(* IEC 61131-3 sources: plc-st-coding-agent/progress/evidence/f14_v14_remaining_20261113/jobs/custom_minimax-m27 (part 2) *)

(* ---- public-hard-03.raw_candidate_01.st ---- *)
FUNCTION_BLOCK FB_RecipeManager
VAR_INPUT
    addRecipe      : BOOL;
    deleteRecipe   : BOOL;
    modifyRecipe   : BOOL;
    queryRecipe    : BOOL;
    recipeIn       : ST_Recipe;
END_VAR

VAR_OUTPUT
    recipeAdded        : BOOL;
    recipeDeleted      : BOOL;
    recipeModified     : BOOL;
    recipeQueryResult  : ST_Recipe;
    error              : BOOL;
    status             : WORD;
END_VAR

VAR_IN_OUT
    recipe : ARRAY[1..10] OF ST_Recipe;
END_VAR

VAR
    tmp_foundIndex : INT;
    tmp_emptyIndex : INT;
    tmp_i          : INT;
END_VAR

(*
ENGINEERING_CONTRACT
===================
Operation sequencing (PUB001-PUB005, PUB007-PUB012):
- Commands evaluated in priority order: DELETE > ADD > MODIFY > QUERY when multiple asserted.
- All success pulses are same-scan; no retention across scans.

Query (PUB008):
  Activation:    queryRecipe rising edge or held high during scan.
  Retention:     recipeQueryResult valid until next scan or successful QUERY.
  Reset:         error and status cleared at start of scan.
  Error codes:   16#8001 = recipe not found.
  Units:         Status WORD error code.

Add (PUB009):
  Activation:    addRecipe rising edge or held high.
  Retention:     Stored in smallest-index empty slot; persists until delete.
  Reset:         None (persistent storage).
  Error codes:   16#8002 = duplicate ID; 16#8003 = database full.
  Same-scan:     Duplicate check before empty-slot check.

Delete (PUB010):
  Activation:    deleteRecipe rising edge or held high.
  Retention:     recipeID forced to 0 (empty slot marker).
  Reset:         Implicit (setting ID to 0 removes it).
  Error codes:   16#8004 = recipe not found.

Modify (PUB011-PUB012):
  Activation:    modifyRecipe rising edge or held high.
  Retention:     Full recipe replacement at found slot.
  Reset:         None.
  Error codes:   16#8005 = recipe not found.
*)

(* CONTRACT_RULES [] *)

tmp_foundIndex := 0;
tmp_emptyIndex := 0;
error := FALSE;
status := 16#0;
recipeAdded := FALSE;
recipeDeleted := FALSE;
recipeModified := FALSE;

IF deleteRecipe THEN
    tmp_foundIndex := 0;
    FOR tmp_i := 1 TO 10 DO
        IF recipe[tmp_i].recipeID <> 0 AND recipe[tmp_i].recipeID = recipeIn.recipeID THEN
            tmp_foundIndex := tmp_i;
            EXIT;
        END_IF
    END_FOR;

    IF tmp_foundIndex = 0 THEN
        error := TRUE;
        status := 16#8004;
    ELSE
        recipe[tmp_foundIndex].recipeID := 0;
        recipeDeleted := TRUE;
    END_IF;

ELSIF addRecipe THEN
    tmp_foundIndex := 0;
    tmp_emptyIndex := 0;

    FOR tmp_i := 1 TO 10 DO
        IF recipe[tmp_i].recipeID <> 0 AND recipe[tmp_i].recipeID = recipeIn.recipeID THEN
            tmp_foundIndex := tmp_i;
            EXIT;
        END_IF
    END_FOR;

    IF tmp_foundIndex <> 0 THEN
        error := TRUE;
        status := 16#8002;
    ELSE
        FOR tmp_i := 1 TO 10 DO
            IF recipe[tmp_i].recipeID = 0 AND tmp_emptyIndex = 0 THEN
                tmp_emptyIndex := tmp_i;
                EXIT;
            END_IF
        END_FOR;

        IF tmp_emptyIndex = 0 THEN
            error := TRUE;
            status := 16#8003;
        ELSE
            recipe[tmp_emptyIndex] := recipeIn;
            recipeAdded := TRUE;
        END_IF;
    END_IF;

ELSIF modifyRecipe THEN
    tmp_foundIndex := 0;
    FOR tmp_i := 1 TO 10 DO
        IF recipe[tmp_i].recipeID <> 0 AND recipe[tmp_i].recipeID = recipeIn.recipeID THEN
            tmp_foundIndex := tmp_i;
            EXIT;
        END_IF
    END_FOR;

    IF tmp_foundIndex = 0 THEN
        error := TRUE;
        status := 16#8005;
    ELSE
        recipe[tmp_foundIndex] := recipeIn;
        recipeModified := TRUE;
    END_IF;

ELSIF queryRecipe THEN
    tmp_foundIndex := 0;
    FOR tmp_i := 1 TO 10 DO
        IF recipe[tmp_i].recipeID <> 0 AND recipe[tmp_i].recipeID = recipeIn.recipeID THEN
            tmp_foundIndex := tmp_i;
            EXIT;
        END_IF
    END_FOR;

    IF tmp_foundIndex = 0 THEN
        error := TRUE;
        status := 16#8001;
    ELSE
        recipeQueryResult := recipe[tmp_foundIndex];
    END_IF;
END_IF;

END_FUNCTION_BLOCK

(* ---- public-hard-03.raw_candidate_02.st ---- *)
TYPE ST_Recipe :
STRUCT
    recipeID               : INT;
    ingredientType         : INT;
    ingredientRatio        : REAL;
    productionTemperature  : REAL;
END_STRUCT
END_TYPE

FUNCTION_BLOCK FB_RecipeManager
VAR_INPUT
    addRecipe      : BOOL;
    deleteRecipe   : BOOL;
    modifyRecipe   : BOOL;
    queryRecipe    : BOOL;
    recipeIn       : ST_Recipe;
END_VAR

VAR_OUTPUT
    recipeAdded        : BOOL;
    recipeDeleted      : BOOL;
    recipeModified     : BOOL;
    recipeQueryResult  : ST_Recipe;
    error              : BOOL;
    status             : WORD;
END_VAR

VAR_IN_OUT
    recipe : ARRAY[1..10] OF ST_Recipe;
END_VAR

VAR
    tmp_foundIndex : INT;
    tmp_emptyIndex : INT;
    tmp_i          : INT;
END_VAR

(*
ENGINEERING_CONTRACT
===================
Operation sequencing (PUB001-PUB005, PUB007-PUB012):
- Commands evaluated in priority order: DELETE > ADD > MODIFY > QUERY when multiple asserted.
- All success pulses are same-scan; no retention across scans.

Query (PUB008):
  Activation:    queryRecipe rising edge or held high during scan.
  Retention:     recipeQueryResult valid until next scan or successful QUERY.
  Reset:         error and status cleared at start of scan.
  Error codes:   16#8001 = recipe not found.
  Units:         Status WORD error code.

Add (PUB009):
  Activation:    addRecipe rising edge or held high.
  Retention:     Stored in smallest-index empty slot; persists until delete.
  Reset:         None (persistent storage).
  Error codes:   16#8002 = duplicate ID; 16#8003 = database full.
  Same-scan:     Duplicate check before empty-slot check.

Delete (PUB010):
  Activation:    deleteRecipe rising edge or held high.
  Retention:     recipeID forced to 0 (empty slot marker).
  Reset:         Implicit (setting ID to 0 removes it).
  Error codes:   16#8004 = recipe not found.

Modify (PUB011-PUB012):
  Activation:    modifyRecipe rising edge or held high.
  Retention:     Full recipe replacement at found slot.
  Reset:         None.
  Error codes:   16#8005 = recipe not found.
*)

(* CONTRACT_RULES [] *)

tmp_foundIndex := 0;
tmp_emptyIndex := 0;
error := FALSE;
status := 16#0;
recipeAdded := FALSE;
recipeDeleted := FALSE;
recipeModified := FALSE;

IF deleteRecipe THEN
    tmp_foundIndex := 0;
    FOR tmp_i := 1 TO 10 DO
        IF recipe[tmp_i].recipeID <> 0 AND recipe[tmp_i].recipeID = recipeIn.recipeID THEN
            tmp_foundIndex := tmp_i;
            EXIT;
        END_IF;
    END_FOR;

    IF tmp_foundIndex = 0 THEN
        error := TRUE;
        status := 16#8004;
    ELSE
        recipe[tmp_foundIndex].recipeID := 0;
        recipeDeleted := TRUE;
    END_IF;

ELSIF addRecipe THEN
    tmp_foundIndex := 0;
    tmp_emptyIndex := 0;

    FOR tmp_i := 1 TO 10 DO
        IF recipe[tmp_i].recipeID <> 0 AND recipe[tmp_i].recipeID = recipeIn.recipeID THEN
            tmp_foundIndex := tmp_i;
            EXIT;
        END_IF;
    END_FOR;

    IF tmp_foundIndex <> 0 THEN
        error := TRUE;
        status := 16#8002;
    ELSE
        FOR tmp_i := 1 TO 10 DO
            IF recipe[tmp_i].recipeID = 0 AND tmp_emptyIndex = 0 THEN
                tmp_emptyIndex := tmp_i;
                EXIT;
            END_IF;
        END_FOR;

        IF tmp_emptyIndex = 0 THEN
            error := TRUE;
            status := 16#8003;
        ELSE
            recipe[tmp_emptyIndex] := recipeIn;
            recipeAdded := TRUE;
        END_IF;
    END_IF;

ELSIF modifyRecipe THEN
    tmp_foundIndex := 0;
    FOR tmp_i := 1 TO 10 DO
        IF recipe[tmp_i].recipeID <> 0 AND recipe[tmp_i].recipeID = recipeIn.recipeID THEN
            tmp_foundIndex := tmp_i;
            EXIT;
        END_IF;
    END_FOR;

    IF tmp_foundIndex = 0 THEN
        error := TRUE;
        status := 16#8005;
    ELSE
        recipe[tmp_foundIndex] := recipeIn;
        recipeModified := TRUE;
    END_IF;

ELSIF queryRecipe THEN
    tmp_foundIndex := 0;
    FOR tmp_i := 1 TO 10 DO
        IF recipe[tmp_i].recipeID <> 0 AND recipe[tmp_i].recipeID = recipeIn.recipeID THEN
            tmp_foundIndex := tmp_i;
            EXIT;
        END_IF;
    END_FOR;

    IF tmp_foundIndex = 0 THEN
        error := TRUE;
        status := 16#8001;
    ELSE
        recipeQueryResult := recipe[tmp_foundIndex];
    END_IF;
END_IF;

END_FUNCTION_BLOCK

(* ---- public-hard-04.candidate_01.st ---- *)
FUNCTION_BLOCK FB
VAR_INPUT
    enqueue  : BOOL;
    dequeue  : BOOL;
    reset    : BOOL;
END_VAR
VAR_OUTPUT
    elementCount : DINT := 0;
    status       : WORD := 16#0000;
END_VAR
VAR_IN_OUT
    item   : VARIANT;
    buffer : VARIANT;
END_VAR
VAR
    head          : DINT := 0;
    tail          : DINT := 0;
    enqueue_prev  : BOOL := FALSE;
    dequeue_prev  : BOOL := FALSE;
    enqueue_trig  : R_TRIG;
    dequeue_trig  : R_TRIG;
    tmp_lower     : DINT;
    tmp_upper     : DINT;
    tmp_capacity  : DINT;
    tmp_element   : DINT;
END_VAR
VAR_TEMP
    emptyArray : ARRAY[0..0] OF DINT;
END_VAR
// ENGINEERING_CONTRACT
// ─────────────────────────────────────────────────────────────────────────────
// PUB001: enqueue rising edge → write item to tail; reject if elementCount == capacity.
// PUB002: dequeue rising edge → read buffer[head] to item; reject if elementCount == 0.
// PUB003: reset TRUE → head:=0, tail:=0, elementCount:=0; no buffer overwrite.
// PUB004: elementCount output tracks live queue size (0..capacity).
// PUB005: status 16#0000=no error/idle; 16#8001=dequeue reject (empty);
//         16#8002=enqueue reject (full); 16#8003=simultaneous enqueue+dequeue.
// PUB006: buffer is caller-supplied VARIANT array; capacity = UPPER-LOWER+1.
// PUB007: item is VARIANT scalar; type must match buffer element type.
// PUB008: circular queue uses head (read index) and tail (write index) modulo capacity.
// PUB009: first invocation initializes to empty state (no prior buffer content used).
// PUB010: reset has priority over enqueue/dequeue.
// PUB011: simultaneous enqueue+dequeue is invalid usage → rejected with status 16#8003.
// ─────────────────────────────────────────────────────────────────────────────
// (* CONTRACT_RULES [] *)
// ─────────────────────────────────────────────────────────────────────────────
    // Capture rising edges for enqueue and dequeue commands
    enqueue_trig(CLK := enqueue);
    dequeue_trig(CLK := dequeue);

    // Update previous state for next scan edge detection
    enqueue_prev  := enqueue;
    dequeue_prev  := dequeue;

    // Reject simultaneous enqueue and dequeue requests
    IF enqueue AND dequeue THEN
        status := 16#8003;
        RETURN;
    END_IF;

    // Validate buffer pointer and extract array bounds
    IF __ISVALIDPTR(buffer, TO_DINT(SIZEOF(emptyArray))) THEN
        tmp_lower    := LOWER_BOUND(buffer, 1);
        tmp_upper    := UPPER_BOUND(buffer, 1);
        tmp_capacity := TO_DINT(tmp_upper - tmp_lower + 1);

        // Validate capacity is positive
        IF tmp_capacity <= 0 THEN
            status := 16#FFFF;
            RETURN;
        END_IF;

        // Type validation: ensure item type matches buffer element type
        // by reading from buffer then assigning to item (runtime type check)
        tmp_element := buffer[tmp_lower];
        tmp_element := item;

        // Execute prioritized operations
        IF reset THEN
            // PUB003: Reset clears queue state without overwriting buffer content
            head        := 0;
            tail        := 0;
            elementCount := 0;
            status      := 16#0000;
        ELSIF enqueue_trig.Q THEN
            // PUB001: Enqueue operation
            IF elementCount >= tmp_capacity THEN
                // Queue full - reject enqueue
                status := 16#8002;
            ELSE
                // Write item to tail position, advance tail circularly
                buffer[tail] := item;
                tail         := (tail + 1) MOD tmp_capacity;
                elementCount := elementCount + 1;
                status       := 16#0000;
            END_IF;
        ELSIF dequeue_trig.Q THEN
            // PUB002: Dequeue operation
            IF elementCount <= 0 THEN
                // Queue empty - reject dequeue
                status := 16#8001;
            ELSE
                // Read from head position, advance head circularly
                item        := buffer[head];
                head        := (head + 1) MOD tmp_capacity;
                elementCount := elementCount - 1;
                status       := 16#0000;
            END_IF;
        ELSE
            // No operation requested this scan
            status := 16#0000;
        END_IF;
    ELSE
        status := 16#FFFF;
    END_IF;
END_FUNCTION_BLOCK

(* ---- public-hard-04.candidate_03.st ---- *)
FUNCTION_BLOCK FB
VAR_INPUT
    enqueue  : BOOL;
    dequeue  : BOOL;
    reset    : BOOL;
END_VAR
VAR_OUTPUT
    elementCount : DINT := 0;
    status       : WORD := 16#0000;
END_VAR
VAR_IN_OUT
    item   : VARIANT;
    buffer : VARIANT;
END_VAR
VAR
    head          : DINT := 0;
    tail          : DINT := 0;
    enqueue_prev  : BOOL := FALSE;
    dequeue_prev  : BOOL := FALSE;
    enqueue_trig  : R_TRIG;
    dequeue_trig  : R_TRIG;
    tmp_lower     : DINT;
    tmp_upper     : DINT;
    tmp_capacity  : DINT;
    tmp_element   : DINT;
END_VAR
// ENGINEERING_CONTRACT
// ─────────────────────────────────────────────────────────────────────────────
// PUB001: enqueue rising edge → write item to tail; reject if elementCount == capacity.
// PUB002: dequeue rising edge → read buffer[head] to item; reject if elementCount == 0.
// PUB003: reset TRUE → head:=0, tail:=0, elementCount:=0; no buffer overwrite.
// PUB004: elementCount output tracks live queue size (0..capacity).
// PUB005: status 16#0000=no error/idle; 16#8001=dequeue reject (empty);
//         16#8002=enqueue reject (full); 16#8003=simultaneous enqueue+dequeue.
// PUB006: buffer is caller-supplied VARIANT array; capacity = UPPER-LOWER+1.
// PUB007: item is VARIANT scalar; type must match buffer element type.
// PUB008: circular queue uses head (read index) and tail (write index) modulo capacity.
// PUB009: first invocation initializes to empty state (no prior buffer content used).
// PUB010: reset has priority over enqueue/dequeue.
// PUB011: simultaneous enqueue+dequeue is invalid usage → rejected with status 16#8003.
// ─────────────────────────────────────────────────────────────────────────────
// (* CONTRACT_RULES [] *)
// ─────────────────────────────────────────────────────────────────────────────
    // Capture rising edges for enqueue and dequeue commands
    enqueue_trig(CLK := enqueue);
    dequeue_trig(CLK := dequeue);

    // Reject simultaneous enqueue and dequeue requests
    IF enqueue AND dequeue THEN
        status := 16#8003;
        RETURN;
    END_IF;

    // Extract array bounds from caller-supplied buffer
    tmp_lower    := LOWER_BOUND(buffer, 1);
    tmp_upper    := UPPER_BOUND(buffer, 1);
    tmp_capacity := tmp_upper - tmp_lower + 1;

    // Execute prioritized operations
    IF reset THEN
        // PUB003: Reset clears queue state without overwriting buffer content
        head         := 0;
        tail         := 0;
        elementCount := 0;
        status       := 16#0000;
    ELSIF enqueue_trig.Q THEN
        // PUB001: Enqueue operation
        IF elementCount >= tmp_capacity THEN
            // Queue full - reject enqueue
            status := 16#8002;
        ELSE
            // Write item to tail position, advance tail circularly
            buffer[tail] := item;
            tail         := (tail + 1) MOD tmp_capacity;
            elementCount := elementCount + 1;
            status       := 16#0000;
        END_IF;
    ELSIF dequeue_trig.Q THEN
        // PUB002: Dequeue operation
        IF elementCount <= 0 THEN
            // Queue empty - reject dequeue
            status := 16#8001;
        ELSE
            // Read from head position, advance head circularly
            item        := buffer[head];
            head        := (head + 1) MOD tmp_capacity;
            elementCount := elementCount - 1;
            status       := 16#0000;
        END_IF;
    ELSE
        // No operation requested this scan
        status := 16#0000;
    END_IF;
END_FUNCTION_BLOCK

(* ---- public-hard-04.patch_base_02.st ---- *)
FUNCTION_BLOCK FB
VAR_INPUT
    enqueue  : BOOL;
    dequeue  : BOOL;
    reset    : BOOL;
END_VAR
VAR_OUTPUT
    elementCount : DINT := 0;
    status       : WORD := 16#0000;
END_VAR
VAR_IN_OUT
    item   : VARIANT;
    buffer : VARIANT;
END_VAR
VAR
    head          : DINT := 0;
    tail          : DINT := 0;
    enqueue_prev  : BOOL := FALSE;
    dequeue_prev  : BOOL := FALSE;
    enqueue_trig  : R_TRIG;
    dequeue_trig  : R_TRIG;
    tmp_lower     : DINT;
    tmp_upper     : DINT;
    tmp_capacity  : DINT;
    tmp_element   : DINT;
END_VAR
VAR_TEMP
    emptyArray : ARRAY[0..0] OF DINT;
END_VAR
// ENGINEERING_CONTRACT
// ─────────────────────────────────────────────────────────────────────────────
// PUB001: enqueue rising edge → write item to tail; reject if elementCount == capacity.
// PUB002: dequeue rising edge → read buffer[head] to item; reject if elementCount == 0.
// PUB003: reset TRUE → head:=0, tail:=0, elementCount:=0; no buffer overwrite.
// PUB004: elementCount output tracks live queue size (0..capacity).
// PUB005: status 16#0000=no error/idle; 16#8001=dequeue reject (empty);
//         16#8002=enqueue reject (full); 16#8003=simultaneous enqueue+dequeue.
// PUB006: buffer is caller-supplied VARIANT array; capacity = UPPER-LOWER+1.
// PUB007: item is VARIANT scalar; type must match buffer element type.
// PUB008: circular queue uses head (read index) and tail (write index) modulo capacity.
// PUB009: first invocation initializes to empty state (no prior buffer content used).
// PUB010: reset has priority over enqueue/dequeue.
// PUB011: simultaneous enqueue+dequeue is invalid usage → rejected with status 16#8003.
// ─────────────────────────────────────────────────────────────────────────────
// (* CONTRACT_RULES [] *)
// ─────────────────────────────────────────────────────────────────────────────
    // Capture rising edges for enqueue and dequeue commands
    enqueue_trig(CLK := enqueue);
    dequeue_trig(CLK := dequeue);

    // Update previous state for next scan edge detection
    enqueue_prev  := enqueue;
    dequeue_prev  := dequeue;

    // Reject simultaneous enqueue and dequeue requests
    IF enqueue AND dequeue THEN
        status := 16#8003;
        RETURN;
    END_IF;

    // Validate buffer pointer and extract array bounds
    IF __ISVALIDPTR(buffer, TO_DINT(SIZEOF(emptyArray))) THEN
        tmp_lower    := LOWER_BOUND(buffer, 1);
        tmp_upper    := UPPER_BOUND(buffer, 1);
        tmp_capacity := TO_DINT(tmp_upper - tmp_lower + 1);

        // Validate capacity is positive
        IF tmp_capacity <= 0 THEN
            status := 16#FFFF;
            RETURN;
        END_IF;

        // Type validation: ensure item type matches buffer element type
        // by reading from buffer then assigning to item (runtime type check)
        tmp_element := buffer[tmp_lower];
        tmp_element := item;

        // Execute prioritized operations
        IF reset THEN
            // PUB003: Reset clears queue state without overwriting buffer content
            head        := 0;
            tail        := 0;
            elementCount := 0;
            status      := 16#0000;
        ELSIF enqueue_trig.Q THEN
            // PUB001: Enqueue operation
            IF elementCount >= tmp_capacity THEN
                // Queue full - reject enqueue
                status := 16#8002;
            ELSE
                // Write item to tail position, advance tail circularly
                buffer[tail] := item;
                tail         := (tail + 1) MOD tmp_capacity;
                elementCount := elementCount + 1;
                status       := 16#0000;
            END_IF;
        ELSIF dequeue_trig.Q THEN
            // PUB002: Dequeue operation
            IF elementCount <= 0 THEN
                // Queue empty - reject dequeue
                status := 16#8001;
            ELSE
                // Read from head position, advance head circularly
                item        := buffer[head];
                head        := (head + 1) MOD tmp_capacity;
                elementCount := elementCount - 1;
                status       := 16#0000;
            END_IF;
        ELSE
            // No operation requested this scan
            status := 16#0000;
        END_IF;
    ELSE
        status := 16#FFFF;
    END_IF;
END_FUNCTION_BLOCK

(* ---- public-hard-04.patch_base_03.st ---- *)
FUNCTION_BLOCK FB
VAR_INPUT
    enqueue  : BOOL;
    dequeue  : BOOL;
    reset    : BOOL;
END_VAR
VAR_OUTPUT
    elementCount : DINT := 0;
    status       : WORD := 16#0000;
END_VAR
VAR_IN_OUT
    item   : VARIANT;
    buffer : VARIANT;
END_VAR
VAR
    head          : DINT := 0;
    tail          : DINT := 0;
    enqueue_prev  : BOOL := FALSE;
    dequeue_prev  : BOOL := FALSE;
    enqueue_trig  : R_TRIG;
    dequeue_trig  : R_TRIG;
    tmp_lower     : DINT;
    tmp_upper     : DINT;
    tmp_capacity  : DINT;
    tmp_element   : DINT;
END_VAR
VAR_TEMP
    emptyArray : ARRAY[0..0] OF DINT;
END_VAR
// ENGINEERING_CONTRACT
// ─────────────────────────────────────────────────────────────────────────────
// PUB001: enqueue rising edge → write item to tail; reject if elementCount == capacity.
// PUB002: dequeue rising edge → read buffer[head] to item; reject if elementCount == 0.
// PUB003: reset TRUE → head:=0, tail:=0, elementCount:=0; no buffer overwrite.
// PUB004: elementCount output tracks live queue size (0..capacity).
// PUB005: status 16#0000=no error/idle; 16#8001=dequeue reject (empty);
//         16#8002=enqueue reject (full); 16#8003=simultaneous enqueue+dequeue.
// PUB006: buffer is caller-supplied VARIANT array; capacity = UPPER-LOWER+1.
// PUB007: item is VARIANT scalar; type must match buffer element type.
// PUB008: circular queue uses head (read index) and tail (write index) modulo capacity.
// PUB009: first invocation initializes to empty state (no prior buffer content used).
// PUB010: reset has priority over enqueue/dequeue.
// PUB011: simultaneous enqueue+dequeue is invalid usage → rejected with status 16#8003.
// ─────────────────────────────────────────────────────────────────────────────
// (* CONTRACT_RULES [] *)
// ─────────────────────────────────────────────────────────────────────────────
    // Capture rising edges for enqueue and dequeue commands
    enqueue_trig(CLK := enqueue);
    dequeue_trig(CLK := dequeue);

    // Update previous state for next scan edge detection
    enqueue_prev  := enqueue;
    dequeue_prev  := dequeue;

    // Reject simultaneous enqueue and dequeue requests
    IF enqueue AND dequeue THEN
        status := 16#8003;
        RETURN;
    END_IF;

    // Validate buffer pointer and extract array bounds
    IF __ISVALIDPTR(buffer, TO_DINT(SIZEOF(emptyArray))) THEN
        tmp_lower    := LOWER_BOUND(buffer, 1);
        tmp_upper    := UPPER_BOUND(buffer, 1);
        tmp_capacity := TO_DINT(tmp_upper - tmp_lower + 1);

        // Validate capacity is positive
        IF tmp_capacity <= 0 THEN
            status := 16#FFFF;
            RETURN;
        END_IF;

        // Type validation: ensure item type matches buffer element type
        // by reading from buffer then assigning to item (runtime type check)
        tmp_element := buffer[tmp_lower];
        tmp_element := item;

        // Execute prioritized operations
        IF reset THEN
            // PUB003: Reset clears queue state without overwriting buffer content
            head        := 0;
            tail        := 0;
            elementCount := 0;
            status      := 16#0000;
        ELSIF enqueue_trig.Q THEN
            // PUB001: Enqueue operation
            IF elementCount >= tmp_capacity THEN
                // Queue full - reject enqueue
                status := 16#8002;
            ELSE
                // Write item to tail position, advance tail circularly
                buffer[tail] := item;
                tail         := (tail + 1) MOD tmp_capacity;
                elementCount := elementCount + 1;
                status       := 16#0000;
            END_IF;
        ELSIF dequeue_trig.Q THEN
            // PUB002: Dequeue operation
            IF elementCount <= 0 THEN
                // Queue empty - reject dequeue
                status := 16#8001;
            ELSE
                // Read from head position, advance head circularly
                item        := buffer[head];
                head        := (head + 1) MOD tmp_capacity;
                elementCount := elementCount - 1;
                status       := 16#0000;
            END_IF;
        ELSE
            // No operation requested this scan
            status := 16#0000;
        END_IF;
    ELSE
        status := 16#FFFF;
    END_IF;
END_FUNCTION_BLOCK

(* ---- public-hard-04.patch_base_04.st ---- *)
FUNCTION_BLOCK FB
VAR_INPUT
    enqueue  : BOOL;
    dequeue  : BOOL;
    reset    : BOOL;
END_VAR
VAR_OUTPUT
    elementCount : DINT := 0;
    status       : WORD := 16#0000;
END_VAR
VAR_IN_OUT
    item   : VARIANT;
    buffer : VARIANT;
END_VAR
VAR
    head          : DINT := 0;
    tail          : DINT := 0;
    enqueue_prev  : BOOL := FALSE;
    dequeue_prev  : BOOL := FALSE;
    enqueue_trig  : R_TRIG;
    dequeue_trig  : R_TRIG;
    tmp_lower     : DINT;
    tmp_upper     : DINT;
    tmp_capacity  : DINT;
    tmp_element   : DINT;
END_VAR
// ENGINEERING_CONTRACT
// ─────────────────────────────────────────────────────────────────────────────
// PUB001: enqueue rising edge → write item to tail; reject if elementCount == capacity.
// PUB002: dequeue rising edge → read buffer[head] to item; reject if elementCount == 0.
// PUB003: reset TRUE → head:=0, tail:=0, elementCount:=0; no buffer overwrite.
// PUB004: elementCount output tracks live queue size (0..capacity).
// PUB005: status 16#0000=no error/idle; 16#8001=dequeue reject (empty);
//         16#8002=enqueue reject (full); 16#8003=simultaneous enqueue+dequeue.
// PUB006: buffer is caller-supplied VARIANT array; capacity = UPPER-LOWER+1.
// PUB007: item is VARIANT scalar; type must match buffer element type.
// PUB008: circular queue uses head (read index) and tail (write index) modulo capacity.
// PUB009: first invocation initializes to empty state (no prior buffer content used).
// PUB010: reset has priority over enqueue/dequeue.
// PUB011: simultaneous enqueue+dequeue is invalid usage → rejected with status 16#8003.
// ─────────────────────────────────────────────────────────────────────────────
// (* CONTRACT_RULES [] *)
// ─────────────────────────────────────────────────────────────────────────────
    // Capture rising edges for enqueue and dequeue commands
    enqueue_trig(CLK := enqueue);
    dequeue_trig(CLK := dequeue);

    // Reject simultaneous enqueue and dequeue requests
    IF enqueue AND dequeue THEN
        status := 16#8003;
        RETURN;
    END_IF;

    // Extract array bounds from caller-supplied buffer
    tmp_lower    := LOWER_BOUND(buffer, 1);
    tmp_upper    := UPPER_BOUND(buffer, 1);
    tmp_capacity := tmp_upper - tmp_lower + 1;

    // Execute prioritized operations
    IF reset THEN
        // PUB003: Reset clears queue state without overwriting buffer content
        head         := 0;
        tail         := 0;
        elementCount := 0;
        status       := 16#0000;
    ELSIF enqueue_trig.Q THEN
        // PUB001: Enqueue operation
        IF elementCount >= tmp_capacity THEN
            // Queue full - reject enqueue
            status := 16#8002;
        ELSE
            // Write item to tail position, advance tail circularly
            buffer[tail] := item;
            tail         := (tail + 1) MOD tmp_capacity;
            elementCount := elementCount + 1;
            status       := 16#0000;
        END_IF;
    ELSIF dequeue_trig.Q THEN
        // PUB002: Dequeue operation
        IF elementCount <= 0 THEN
            // Queue empty - reject dequeue
            status := 16#8001;
        ELSE
            // Read from head position, advance head circularly
            item        := buffer[head];
            head        := (head + 1) MOD tmp_capacity;
            elementCount := elementCount - 1;
            status       := 16#0000;
        END_IF;
    ELSE
        // No operation requested this scan
        status := 16#0000;
    END_IF;
END_FUNCTION_BLOCK

(* ---- public-hard-04.raw_candidate_01.st ---- *)
FUNCTION_BLOCK FB
VAR_INPUT
    enqueue  : BOOL;
    dequeue  : BOOL;
    reset    : BOOL;
END_VAR
VAR_OUTPUT
    elementCount : DINT := 0;
    status       : WORD := 16#0000;
END_VAR
VAR_IN_OUT
    item   : VARIANT;
    buffer : VARIANT;
END_VAR
VAR
    head          : DINT := 0;
    tail          : DINT := 0;
    enqueue_prev  : BOOL := FALSE;
    dequeue_prev  : BOOL := FALSE;
    enqueue_trig  : R_TRIG;
    dequeue_trig  : R_TRIG;
    tmp_lower     : DINT;
    tmp_upper     : DINT;
    tmp_capacity  : DINT;
    tmp_element   : DINT;
END_VAR
VAR_TEMP
    emptyArray : ARRAY[0..0] OF DINT;
END_VAR
// ENGINEERING_CONTRACT
// ─────────────────────────────────────────────────────────────────────────────
// PUB001: enqueue rising edge → write item to tail; reject if elementCount == capacity.
// PUB002: dequeue rising edge → read buffer[head] to item; reject if elementCount == 0.
// PUB003: reset TRUE → head:=0, tail:=0, elementCount:=0; no buffer overwrite.
// PUB004: elementCount output tracks live queue size (0..capacity).
// PUB005: status 16#0000=no error/idle; 16#8001=dequeue reject (empty);
//         16#8002=enqueue reject (full); 16#8003=simultaneous enqueue+dequeue.
// PUB006: buffer is caller-supplied VARIANT array; capacity = UPPER-LOWER+1.
// PUB007: item is VARIANT scalar; type must match buffer element type.
// PUB008: circular queue uses head (read index) and tail (write index) modulo capacity.
// PUB009: first invocation initializes to empty state (no prior buffer content used).
// PUB010: reset has priority over enqueue/dequeue.
// PUB011: simultaneous enqueue+dequeue is invalid usage → rejected with status 16#8003.
// ─────────────────────────────────────────────────────────────────────────────
// (* CONTRACT_RULES [] *)
// ─────────────────────────────────────────────────────────────────────────────
    // Capture rising edges for enqueue and dequeue commands
    enqueue_trig(CLK := enqueue);
    dequeue_trig(CLK := dequeue);

    // Update previous state for next scan edge detection
    enqueue_prev  := enqueue;
    dequeue_prev  := dequeue;

    // Reject simultaneous enqueue and dequeue requests
    IF enqueue AND dequeue THEN
        status := 16#8003;
        RETURN;
    END_IF

    // Validate buffer pointer and extract array bounds
    IF __ISVALIDPTR(buffer, TO_DINT(SIZEOF(emptyArray))) THEN
        tmp_lower    := LOWER_BOUND(buffer, 1);
        tmp_upper    := UPPER_BOUND(buffer, 1);
        tmp_capacity := TO_DINT(tmp_upper - tmp_lower + 1);

        // Validate capacity is positive
        IF tmp_capacity <= 0 THEN
            status := 16#FFFF;
            RETURN;
        END_IF

        // Type validation: ensure item type matches buffer element type
        // by reading from buffer then assigning to item (runtime type check)
        tmp_element := buffer[tmp_lower];
        tmp_element := item;

        // Execute prioritized operations
        IF reset THEN
            // PUB003: Reset clears queue state without overwriting buffer content
            head        := 0;
            tail        := 0;
            elementCount := 0;
            status      := 16#0000;
        ELSIF enqueue_trig.Q THEN
            // PUB001: Enqueue operation
            IF elementCount >= tmp_capacity THEN
                // Queue full - reject enqueue
                status := 16#8002;
            ELSE
                // Write item to tail position, advance tail circularly
                buffer[tail] := item;
                tail         := (tail + 1) MOD tmp_capacity;
                elementCount := elementCount + 1;
                status       := 16#0000;
            END_IF;
        ELSIF dequeue_trig.Q THEN
            // PUB002: Dequeue operation
            IF elementCount <= 0 THEN
                // Queue empty - reject dequeue
                status := 16#8001;
            ELSE
                // Read from head position, advance head circularly
                item        := buffer[head];
                head        := (head + 1) MOD tmp_capacity;
                elementCount := elementCount - 1;
                status       := 16#0000;
            END_IF;
        ELSE
            // No operation requested this scan
            status := 16#0000;
        END_IF;
    ELSE
        status := 16#FFFF;
    END_IF;
END_FUNCTION_BLOCK

(* ---- public-hard-04.raw_candidate_03.st ---- *)
FUNCTION_BLOCK FB
VAR_INPUT
    enqueue  : BOOL;
    dequeue  : BOOL;
    reset    : BOOL;
END_VAR
VAR_OUTPUT
    elementCount : DINT := 0;
    status       : WORD := 16#0000;
END_VAR
VAR_IN_OUT
    item   : VARIANT;
    buffer : VARIANT;
END_VAR
VAR
    head          : DINT := 0;
    tail          : DINT := 0;
    enqueue_prev  : BOOL := FALSE;
    dequeue_prev  : BOOL := FALSE;
    enqueue_trig  : R_TRIG;
    dequeue_trig  : R_TRIG;
    tmp_lower     : DINT;
    tmp_upper     : DINT;
    tmp_capacity  : DINT;
    tmp_element   : DINT;
END_VAR
// ENGINEERING_CONTRACT
// ─────────────────────────────────────────────────────────────────────────────
// PUB001: enqueue rising edge → write item to tail; reject if elementCount == capacity.
// PUB002: dequeue rising edge → read buffer[head] to item; reject if elementCount == 0.
// PUB003: reset TRUE → head:=0, tail:=0, elementCount:=0; no buffer overwrite.
// PUB004: elementCount output tracks live queue size (0..capacity).
// PUB005: status 16#0000=no error/idle; 16#8001=dequeue reject (empty);
//         16#8002=enqueue reject (full); 16#8003=simultaneous enqueue+dequeue.
// PUB006: buffer is caller-supplied VARIANT array; capacity = UPPER-LOWER+1.
// PUB007: item is VARIANT scalar; type must match buffer element type.
// PUB008: circular queue uses head (read index) and tail (write index) modulo capacity.
// PUB009: first invocation initializes to empty state (no prior buffer content used).
// PUB010: reset has priority over enqueue/dequeue.
// PUB011: simultaneous enqueue+dequeue is invalid usage → rejected with status 16#8003.
// ─────────────────────────────────────────────────────────────────────────────
// (* CONTRACT_RULES [] *)
// ─────────────────────────────────────────────────────────────────────────────
    // Capture rising edges for enqueue and dequeue commands
    enqueue_trig(CLK := enqueue);
    dequeue_trig(CLK := dequeue);

    // Reject simultaneous enqueue and dequeue requests
    IF enqueue AND dequeue THEN
        status := 16#8003;
        RETURN;
    END_IF;

    // Extract array bounds from caller-supplied buffer
    tmp_lower    := LOWER_BOUND(buffer, 1);
    tmp_upper    := UPPER_BOUND(buffer, 1);
    tmp_capacity := tmp_upper - tmp_lower + 1;

    // Execute prioritized operations
    IF reset THEN
        // PUB003: Reset clears queue state without overwriting buffer content
        head         := 0;
        tail         := 0;
        elementCount := 0;
        status       := 16#0000;
    ELSIF enqueue_trig.Q THEN
        // PUB001: Enqueue operation
        IF elementCount >= tmp_capacity THEN
            // Queue full - reject enqueue
            status := 16#8002;
        ELSE
            // Write item to tail position, advance tail circularly
            buffer[tail] := item;
            tail         := (tail + 1) MOD tmp_capacity;
            elementCount := elementCount + 1;
            status       := 16#0000;
        END_IF;
    ELSIF dequeue_trig.Q THEN
        // PUB002: Dequeue operation
        IF elementCount <= 0 THEN
            // Queue empty - reject dequeue
            status := 16#8001;
        ELSE
            // Read from head position, advance head circularly
            item        := buffer[head];
            head        := (head + 1) MOD tmp_capacity;
            elementCount := elementCount - 1;
            status       := 16#0000;
        END_IF;
    ELSE
        // No operation requested this scan
        status := 16#0000;
    END_IF;
END_FUNCTION_BLOCK

(* ---- public-hard-05.candidate_01.st ---- *)
(* ENGINEERING_CONTRACT - Mechanical Arm Control
 * =============================================================================
 * Mode Selection: Caller ensures exactly one mode active; emergency stop has highest priority.
 *
 * Output State Table:
 * | Output          | Activation                              | Retention                     | Reset                        | Priority    |
 * |-----------------|-----------------------------------------|-------------------------------|--------------------------------|-------------|
 * | MoveDown        | Manual:DownButton AND NOT DownLimitSwitch| Manual:button hold; Auto:step | EmergencyStop, step change   | Physical dir |
 * |                 | Auto: current step = down step           | Auto: hold until limit        | button release (manual)       | rule applies |
 * | MoveUp          | Manual:UpButton AND NOT UpLimitSwitch    | Manual:button hold; Auto:step | EmergencyStop, step change   | Physical dir |
 * |                 | Auto: current step = up step             | Auto: hold until limit        | button release (manual)       | rule applies |
 * | MoveLeft        | Manual:LeftButton AND NOT LeftLimitSwitch| Manual:button hold; Auto:step | EmergencyStop, step change   | Physical dir |
 * |                 | Auto: current step = left step           | Auto: hold until limit        | button release (manual)       | rule applies |
 * | MoveRight       | Manual:RightButton AND NOT RightLimitSwitch| Manual:button hold; Auto:step| EmergencyStop, step change   | Physical dir |
 * |                 | Auto: current step = right step          | Auto: hold until limit        | button release (manual)       | rule applies |
 * | ActivateGrip    | Manual:GripButton AND NOT GripLimitSwitch| Manual:button hold; Auto:step | EmergencyStop, step change   | N/A         |
 * |                 | Auto: grip step, hold until GripLimitSwitch| Auto: hold until limit       | button release (manual)       |             |
 * | ActivateRelease | Manual:ReleaseButton AND NOT ReleaseLimitSwitch| Manual:button hold; Auto:step| EmergencyStop, step change  | N/A         |
 * |                 | Auto: release step, hold until ReleaseLimitSwitch| Auto: hold until limit    | button release (manual)       |             |
 *
 * Sequence (8 steps, single cycle and continuous modes):
 *   0: Down -> 1: Grip -> 2: Up -> 3: Right -> 4: Down -> 5: Release -> 6: Up -> 7: Left -> (repeat)
 *
 * Single step mode: Same 8-step sequence, advancing one step per Start rising edge.
 * Single cycle mode: Executes all 8 steps, stops at stepIndex=8.
 * Continuous mode: Executes all 8 steps, returns to stepIndex=0 when complete.
 *
 * Units: Limit switches TRUE=at position (normally-open, closed at position).
 * Boundary: stepIndex ∈ [0..8]; 8 = cycle complete state for single cycle mode.
 * Same-scan: Final output evaluated from current stepIndex and limit switches per scan.
 *
 * Contract PUB clauses: PUB001-PUB020 define all behavior above.
 *)

FUNCTION_BLOCK ArmController
VAR
    stepIndex : INT := 0;         // Current step in sequence (0-7), 8 = single cycle complete
    startButtonPrev : BOOL := FALSE; // Rising edge detection for Start button
    tmpRisingEdge : BOOL;
END_VAR

(* CONTRACT_RULES
[
  {"kind": "hold_until_reset", "output": "MoveDown", "set_input": "DownButton", "reset_input": null},
  {"kind": "hold_until_reset", "output": "MoveUp", "set_input": "UpButton", "reset_input": null},
  {"kind": "hold_until_reset", "output": "MoveLeft", "set_input": "LeftButton", "reset_input": null},
  {"kind": "hold_until_reset", "output": "MoveRight", "set_input": "RightButton", "reset_input": null},
  {"kind": "hold_until_reset", "output": "ActivateGrip", "set_input": "GripButton", "reset_input": null},
  {"kind": "hold_until_reset", "output": "ActivateRelease", "set_input": "ReleaseButton", "reset_input": null}
]
*)

    // Emergency stop has highest priority - stops all outputs
    IF EmergencyStop = FALSE THEN
        MoveDown := FALSE;
        MoveUp := FALSE;
        MoveLeft := FALSE;
        MoveRight := FALSE;
        ActivateGrip := FALSE;
        ActivateRelease := FALSE;
    ELSIF SingleStepMode THEN
        // Detect rising edge on Start button
        tmpRisingEdge := Start AND NOT startButtonPrev;
        startButtonPrev := Start;

        IF tmpRisingEdge THEN
            stepIndex := stepIndex + 1;
            IF stepIndex > 7 THEN
                stepIndex := 0;
            END_IF;
        END_IF;

        // Execute current step
        CASE stepIndex OF
            0: // Down
                MoveDown := TRUE;
                IF DownLimitSwitch THEN
                    stepIndex := 1;
                END_IF;
            1: // Grip
                ActivateGrip := TRUE;
                IF GripLimitSwitch THEN
                    stepIndex := 2;
                END_IF;
            2: // Up
                MoveUp := TRUE;
                IF UpLimitSwitch THEN
                    stepIndex := 3;
                END_IF;
            3: // Right
                MoveRight := TRUE;
                IF RightLimitSwitch THEN
                    stepIndex := 4;
                END_IF;
            4: // Down (second descent)
                MoveDown := TRUE;
                IF DownLimitSwitch THEN
                    stepIndex := 5;
                END_IF;
            5: // Release
                ActivateRelease := TRUE;
                IF ReleaseLimitSwitch THEN
                    stepIndex := 6;
                END_IF;
            6: // Up (second ascent)
                MoveUp := TRUE;
                IF UpLimitSwitch THEN
                    stepIndex := 7;
                END_IF;
            7: // Left (return to start)
                MoveLeft := TRUE;
                IF LeftLimitSwitch THEN
                    stepIndex := 0;
                END_IF;
        END_CASE;

    ELSIF SingleCycleMode THEN
        // Single cycle mode: run through all steps automatically, stop at end
        CASE stepIndex OF
            0:
                MoveDown := NOT DownLimitSwitch;
                IF DownLimitSwitch THEN
                    stepIndex := 1;
                END_IF;
            1:
                ActivateGrip := NOT GripLimitSwitch;
                IF GripLimitSwitch THEN
                    stepIndex := 2;
                END_IF;
            2:
                MoveUp := NOT UpLimitSwitch;
                IF UpLimitSwitch THEN
                    stepIndex := 3;
                END_IF;
            3:
                MoveRight := NOT RightLimitSwitch;
                IF RightLimitSwitch THEN
                    stepIndex := 4;
                END_IF;
            4:
                MoveDown := NOT DownLimitSwitch;
                IF DownLimitSwitch THEN
                    stepIndex := 5;
                END_IF;
            5:
                ActivateRelease := NOT ReleaseLimitSwitch;
                IF ReleaseLimitSwitch THEN
                    stepIndex := 6;
                END_IF;
            6:
                MoveUp := NOT UpLimitSwitch;
                IF UpLimitSwitch THEN
                    stepIndex := 7;
                END_IF;
            7:
                MoveLeft := NOT LeftLimitSwitch;
                IF LeftLimitSwitch THEN
                    stepIndex := 8; // Cycle complete, stay here
                END_IF;
        END_CASE;

    ELSIF ContinuousMode THEN
        // Continuous mode: run through all steps automatically, restart at end
        CASE stepIndex OF
            0:
                MoveDown := NOT DownLimitSwitch;
                IF DownLimitSwitch THEN
                    stepIndex := 1;
                END_IF;
            1:
                ActivateGrip := NOT GripLimitSwitch;
                IF GripLimitSwitch THEN
                    stepIndex := 2;
                END_IF;
            2:
                MoveUp := NOT UpLimitSwitch;
                IF UpLimitSwitch THEN
                    stepIndex := 3;
                END_IF;
            3:
                MoveRight := NOT RightLimitSwitch;
                IF RightLimitSwitch THEN
                    stepIndex := 4;
                END_IF;
            4:
                MoveDown := NOT DownLimitSwitch;
                IF DownLimitSwitch THEN
                    stepIndex := 5;
                END_IF;
            5:
                ActivateRelease := NOT ReleaseLimitSwitch;
                IF ReleaseLimitSwitch THEN
                    stepIndex := 6;
                END_IF;
            6:
                MoveUp := NOT UpLimitSwitch;
                IF UpLimitSwitch THEN
                    stepIndex := 7;
                END_IF;
            7:
                MoveLeft := NOT LeftLimitSwitch;
                IF LeftLimitSwitch THEN
                    stepIndex := 0; // Restart cycle
                END_IF;
        END_CASE;

    ELSIF ManualMode THEN
        // Manual mode: direct button control with limit switch protection
        MoveDown := DownButton AND NOT DownLimitSwitch;
        MoveUp := UpButton AND NOT UpLimitSwitch;
        MoveLeft := LeftButton AND NOT LeftLimitSwitch;
        MoveRight := RightButton AND NOT RightLimitSwitch;
        ActivateGrip := GripButton AND NOT GripLimitSwitch;
        ActivateRelease := ReleaseButton AND NOT ReleaseLimitSwitch;
    END_IF;

END_FUNCTION_BLOCK

(* ---- public-hard-05.candidate_02.st ---- *)
(* ENGINEERING_CONTRACT - Mechanical Arm Control
 * =============================================================================
 * Mode Selection: Caller ensures exactly one mode active; emergency stop has highest priority.
 *
 * Output State Table:
 * | Output          | Activation                              | Retention                     | Reset                        | Priority    |
 * |-----------------|-----------------------------------------|-------------------------------|--------------------------------|-------------|
 * | MoveDown        | Manual:DownButton AND NOT DownLimitSwitch| Manual:button hold; Auto:step | EmergencyStop, step change   | Physical dir |
 * |                 | Auto: current step = down step           | Auto: hold until limit        | button release (manual)       | rule applies |
 * | MoveUp          | Manual:UpButton AND NOT UpLimitSwitch    | Manual:button hold; Auto:step | EmergencyStop, step change   | Physical dir |
 * |                 | Auto: current step = up step             | Auto: hold until limit        | button release (manual)       | rule applies |
 * | MoveLeft        | Manual:LeftButton AND NOT LeftLimitSwitch| Manual:button hold; Auto:step | EmergencyStop, step change   | Physical dir |
 * |                 | Auto: current step = left step           | Auto: hold until limit        | button release (manual)       | rule applies |
 * | MoveRight       | Manual:RightButton AND NOT RightLimitSwitch| Manual:button hold; Auto:step| EmergencyStop, step change   | Physical dir |
 * |                 | Auto: current step = right step          | Auto: hold until limit        | button release (manual)       | rule applies |
 * | ActivateGrip    | Manual:GripButton AND NOT GripLimitSwitch| Manual:button hold; Auto:step | EmergencyStop, step change   | N/A         |
 * |                 | Auto: grip step, hold until GripLimitSwitch| Auto: hold until limit       | button release (manual)       |             |
 * | ActivateRelease | Manual:ReleaseButton AND NOT ReleaseLimitSwitch| Manual:button hold; Auto:step| EmergencyStop, step change  | N/A         |
 * |                 | Auto: release step, hold until ReleaseLimitSwitch| Auto: hold until limit    | button release (manual)       |             |
 *
 * Sequence (8 steps, single cycle and continuous modes):
 *   0: Down -> 1: Grip -> 2: Up -> 3: Right -> 4: Down -> 5: Release -> 6: Up -> 7: Left -> (repeat)
 *
 * Single step mode: Same 8-step sequence, advancing one step per Start rising edge.
 * Single cycle mode: Executes all 8 steps, stops at stepIndex=8.
 * Continuous mode: Executes all 8 steps, returns to stepIndex=0 when complete.
 *
 * Units: Limit switches TRUE=at position (normally-open, closed at position).
 * Boundary: stepIndex ∈ [0..8]; 8 = cycle complete state for single cycle mode.
 * Same-scan: Final output evaluated from current stepIndex and limit switches per scan.
 *
 * Contract PUB clauses: PUB001-PUB020 define all behavior above.
 *)

FUNCTION_BLOCK ArmController
VAR_INPUT
    ManualMode : BOOL;
    SingleStepMode : BOOL;
    SingleCycleMode : BOOL;
    ContinuousMode : BOOL;
    EmergencyStop : BOOL;
    Start : BOOL;
    DownButton : BOOL;
    UpButton : BOOL;
    LeftButton : BOOL;
    RightButton : BOOL;
    GripButton : BOOL;
    ReleaseButton : BOOL;
    DownLimitSwitch : BOOL;
    UpLimitSwitch : BOOL;
    LeftLimitSwitch : BOOL;
    RightLimitSwitch : BOOL;
    GripLimitSwitch : BOOL;
    ReleaseLimitSwitch : BOOL;
END_VAR
VAR_OUTPUT
    MoveDown : BOOL;
    MoveUp : BOOL;
    MoveLeft : BOOL;
    MoveRight : BOOL;
    ActivateGrip : BOOL;
    ActivateRelease : BOOL;
END_VAR
VAR
    stepIndex : INT := 0;         // Current step in sequence (0-7), 8 = single cycle complete
    startButtonPrev : BOOL := FALSE; // Rising edge detection for Start button
    tmpRisingEdge : BOOL;
END_VAR

(* CONTRACT_RULES
[
  {"kind": "hold_until_reset", "output": "MoveDown", "set_input": "DownButton", "reset_input": null},
  {"kind": "hold_until_reset", "output": "MoveUp", "set_input": "UpButton", "reset_input": null},
  {"kind": "hold_until_reset", "output": "MoveLeft", "set_input": "LeftButton", "reset_input": null},
  {"kind": "hold_until_reset", "output": "MoveRight", "set_input": "RightButton", "reset_input": null},
  {"kind": "hold_until_reset", "output": "ActivateGrip", "set_input": "GripButton", "reset_input": null},
  {"kind": "hold_until_reset", "output": "ActivateRelease", "set_input": "ReleaseButton", "reset_input": null}
]
*)

    // Emergency stop has highest priority - stops all outputs
    IF EmergencyStop = FALSE THEN
        MoveDown := FALSE;
        MoveUp := FALSE;
        MoveLeft := FALSE;
        MoveRight := FALSE;
        ActivateGrip := FALSE;
        ActivateRelease := FALSE;
    ELSIF SingleStepMode THEN
        // Detect rising edge on Start button
        tmpRisingEdge := Start AND NOT startButtonPrev;
        startButtonPrev := Start;

        IF tmpRisingEdge THEN
            stepIndex := stepIndex + 1;
            IF stepIndex > 7 THEN
                stepIndex := 0;
            END_IF;
        END_IF;

        // Execute current step
        CASE stepIndex OF
            0: // Down
                MoveDown := TRUE;
                IF DownLimitSwitch THEN
                    stepIndex := 1;
                END_IF;
            1: // Grip
                ActivateGrip := TRUE;
                IF GripLimitSwitch THEN
                    stepIndex := 2;
                END_IF;
            2: // Up
                MoveUp := TRUE;
                IF UpLimitSwitch THEN
                    stepIndex := 3;
                END_IF;
            3: // Right
                MoveRight := TRUE;
                IF RightLimitSwitch THEN
                    stepIndex := 4;
                END_IF;
            4: // Down (second descent)
                MoveDown := TRUE;
                IF DownLimitSwitch THEN
                    stepIndex := 5;
                END_IF;
            5: // Release
                ActivateRelease := TRUE;
                IF ReleaseLimitSwitch THEN
                    stepIndex := 6;
                END_IF;
            6: // Up (second ascent)
                MoveUp := TRUE;
                IF UpLimitSwitch THEN
                    stepIndex := 7;
                END_IF;
            7: // Left (return to start)
                MoveLeft := TRUE;
                IF LeftLimitSwitch THEN
                    stepIndex := 0;
                END_IF;
        END_CASE;

    ELSIF SingleCycleMode THEN
        // Single cycle mode: run through all steps automatically, stop at end
        CASE stepIndex OF
            0:
                MoveDown := NOT DownLimitSwitch;
                IF DownLimitSwitch THEN
                    stepIndex := 1;
                END_IF;
            1:
                ActivateGrip := NOT GripLimitSwitch;
                IF GripLimitSwitch THEN
                    stepIndex := 2;
                END_IF;
            2:
                MoveUp := NOT UpLimitSwitch;
                IF UpLimitSwitch THEN
                    stepIndex := 3;
                END_IF;
            3:
                MoveRight := NOT RightLimitSwitch;
                IF RightLimitSwitch THEN
                    stepIndex := 4;
                END_IF;
            4:
                MoveDown := NOT DownLimitSwitch;
                IF DownLimitSwitch THEN
                    stepIndex := 5;
                END_IF;
            5:
                ActivateRelease := NOT ReleaseLimitSwitch;
                IF ReleaseLimitSwitch THEN
                    stepIndex := 6;
                END_IF;
            6:
                MoveUp := NOT UpLimitSwitch;
                IF UpLimitSwitch THEN
                    stepIndex := 7;
                END_IF;
            7:
                MoveLeft := NOT LeftLimitSwitch;
                IF LeftLimitSwitch THEN
                    stepIndex := 8; // Cycle complete, stay here
                END_IF;
        END_CASE;

    ELSIF ContinuousMode THEN
        // Continuous mode: run through all steps automatically, restart at end
        CASE stepIndex OF
            0:
                MoveDown := NOT DownLimitSwitch;
                IF DownLimitSwitch THEN
                    stepIndex := 1;
                END_IF;
            1:
                ActivateGrip := NOT GripLimitSwitch;
                IF GripLimitSwitch THEN
                    stepIndex := 2;
                END_IF;
            2:
                MoveUp := NOT UpLimitSwitch;
                IF UpLimitSwitch THEN
                    stepIndex := 3;
                END_IF;
            3:
                MoveRight := NOT RightLimitSwitch;
                IF RightLimitSwitch THEN
                    stepIndex := 4;
                END_IF;
            4:
                MoveDown := NOT DownLimitSwitch;
                IF DownLimitSwitch THEN
                    stepIndex := 5;
                END_IF;
            5:
                ActivateRelease := NOT ReleaseLimitSwitch;
                IF ReleaseLimitSwitch THEN
                    stepIndex := 6;
                END_IF;
            6:
                MoveUp := NOT UpLimitSwitch;
                IF UpLimitSwitch THEN
                    stepIndex := 7;
                END_IF;
            7:
                MoveLeft := NOT LeftLimitSwitch;
                IF LeftLimitSwitch THEN
                    stepIndex := 0; // Restart cycle
                END_IF;
        END_CASE;

    ELSIF ManualMode THEN
        // Manual mode: direct button control with limit switch protection
        MoveDown := DownButton AND NOT DownLimitSwitch;
        MoveUp := UpButton AND NOT UpLimitSwitch;
        MoveLeft := LeftButton AND NOT LeftLimitSwitch;
        MoveRight := RightButton AND NOT RightLimitSwitch;
        ActivateGrip := GripButton AND NOT GripLimitSwitch;
        ActivateRelease := ReleaseButton AND NOT ReleaseLimitSwitch;
    END_IF;

END_FUNCTION_BLOCK

(* ---- public-hard-05.patch_base_02.st ---- *)
(* ENGINEERING_CONTRACT - Mechanical Arm Control
 * =============================================================================
 * Mode Selection: Caller ensures exactly one mode active; emergency stop has highest priority.
 *
 * Output State Table:
 * | Output          | Activation                              | Retention                     | Reset                        | Priority    |
 * |-----------------|-----------------------------------------|-------------------------------|--------------------------------|-------------|
 * | MoveDown        | Manual:DownButton AND NOT DownLimitSwitch| Manual:button hold; Auto:step | EmergencyStop, step change   | Physical dir |
 * |                 | Auto: current step = down step           | Auto: hold until limit        | button release (manual)       | rule applies |
 * | MoveUp          | Manual:UpButton AND NOT UpLimitSwitch    | Manual:button hold; Auto:step | EmergencyStop, step change   | Physical dir |
 * |                 | Auto: current step = up step             | Auto: hold until limit        | button release (manual)       | rule applies |
 * | MoveLeft        | Manual:LeftButton AND NOT LeftLimitSwitch| Manual:button hold; Auto:step | EmergencyStop, step change   | Physical dir |
 * |                 | Auto: current step = left step           | Auto: hold until limit        | button release (manual)       | rule applies |
 * | MoveRight       | Manual:RightButton AND NOT RightLimitSwitch| Manual:button hold; Auto:step| EmergencyStop, step change   | Physical dir |
 * |                 | Auto: current step = right step          | Auto: hold until limit        | button release (manual)       | rule applies |
 * | ActivateGrip    | Manual:GripButton AND NOT GripLimitSwitch| Manual:button hold; Auto:step | EmergencyStop, step change   | N/A         |
 * |                 | Auto: grip step, hold until GripLimitSwitch| Auto: hold until limit       | button release (manual)       |             |
 * | ActivateRelease | Manual:ReleaseButton AND NOT ReleaseLimitSwitch| Manual:button hold; Auto:step| EmergencyStop, step change  | N/A         |
 * |                 | Auto: release step, hold until ReleaseLimitSwitch| Auto: hold until limit    | button release (manual)       |             |
 *
 * Sequence (8 steps, single cycle and continuous modes):
 *   0: Down -> 1: Grip -> 2: Up -> 3: Right -> 4: Down -> 5: Release -> 6: Up -> 7: Left -> (repeat)
 *
 * Single step mode: Same 8-step sequence, advancing one step per Start rising edge.
 * Single cycle mode: Executes all 8 steps, stops at stepIndex=8.
 * Continuous mode: Executes all 8 steps, returns to stepIndex=0 when complete.
 *
 * Units: Limit switches TRUE=at position (normally-open, closed at position).
 * Boundary: stepIndex ∈ [0..8]; 8 = cycle complete state for single cycle mode.
 * Same-scan: Final output evaluated from current stepIndex and limit switches per scan.
 *
 * Contract PUB clauses: PUB001-PUB020 define all behavior above.
 *)

FUNCTION_BLOCK ArmController
VAR
    stepIndex : INT := 0;         // Current step in sequence (0-7), 8 = single cycle complete
    startButtonPrev : BOOL := FALSE; // Rising edge detection for Start button
    tmpRisingEdge : BOOL;
END_VAR

(* CONTRACT_RULES
[
  {"kind": "hold_until_reset", "output": "MoveDown", "set_input": "DownButton", "reset_input": null},
  {"kind": "hold_until_reset", "output": "MoveUp", "set_input": "UpButton", "reset_input": null},
  {"kind": "hold_until_reset", "output": "MoveLeft", "set_input": "LeftButton", "reset_input": null},
  {"kind": "hold_until_reset", "output": "MoveRight", "set_input": "RightButton", "reset_input": null},
  {"kind": "hold_until_reset", "output": "ActivateGrip", "set_input": "GripButton", "reset_input": null},
  {"kind": "hold_until_reset", "output": "ActivateRelease", "set_input": "ReleaseButton", "reset_input": null}
]
*)

    // Emergency stop has highest priority - stops all outputs
    IF EmergencyStop = FALSE THEN
        MoveDown := FALSE;
        MoveUp := FALSE;
        MoveLeft := FALSE;
        MoveRight := FALSE;
        ActivateGrip := FALSE;
        ActivateRelease := FALSE;
    ELSIF SingleStepMode THEN
        // Detect rising edge on Start button
        tmpRisingEdge := Start AND NOT startButtonPrev;
        startButtonPrev := Start;

        IF tmpRisingEdge THEN
            stepIndex := stepIndex + 1;
            IF stepIndex > 7 THEN
                stepIndex := 0;
            END_IF;
        END_IF;

        // Execute current step
        CASE stepIndex OF
            0: // Down
                MoveDown := TRUE;
                IF DownLimitSwitch THEN
                    stepIndex := 1;
                END_IF;
            1: // Grip
                ActivateGrip := TRUE;
                IF GripLimitSwitch THEN
                    stepIndex := 2;
                END_IF;
            2: // Up
                MoveUp := TRUE;
                IF UpLimitSwitch THEN
                    stepIndex := 3;
                END_IF;
            3: // Right
                MoveRight := TRUE;
                IF RightLimitSwitch THEN
                    stepIndex := 4;
                END_IF;
            4: // Down (second descent)
                MoveDown := TRUE;
                IF DownLimitSwitch THEN
                    stepIndex := 5;
                END_IF;
            5: // Release
                ActivateRelease := TRUE;
                IF ReleaseLimitSwitch THEN
                    stepIndex := 6;
                END_IF;
            6: // Up (second ascent)
                MoveUp := TRUE;
                IF UpLimitSwitch THEN
                    stepIndex := 7;
                END_IF;
            7: // Left (return to start)
                MoveLeft := TRUE;
                IF LeftLimitSwitch THEN
                    stepIndex := 0;
                END_IF;
        END_CASE;

    ELSIF SingleCycleMode THEN
        // Single cycle mode: run through all steps automatically, stop at end
        CASE stepIndex OF
            0:
                MoveDown := NOT DownLimitSwitch;
                IF DownLimitSwitch THEN
                    stepIndex := 1;
                END_IF;
            1:
                ActivateGrip := NOT GripLimitSwitch;
                IF GripLimitSwitch THEN
                    stepIndex := 2;
                END_IF;
            2:
                MoveUp := NOT UpLimitSwitch;
                IF UpLimitSwitch THEN
                    stepIndex := 3;
                END_IF;
            3:
                MoveRight := NOT RightLimitSwitch;
                IF RightLimitSwitch THEN
                    stepIndex := 4;
                END_IF;
            4:
                MoveDown := NOT DownLimitSwitch;
                IF DownLimitSwitch THEN
                    stepIndex := 5;
                END_IF;
            5:
                ActivateRelease := NOT ReleaseLimitSwitch;
                IF ReleaseLimitSwitch THEN
                    stepIndex := 6;
                END_IF;
            6:
                MoveUp := NOT UpLimitSwitch;
                IF UpLimitSwitch THEN
                    stepIndex := 7;
                END_IF;
            7:
                MoveLeft := NOT LeftLimitSwitch;
                IF LeftLimitSwitch THEN
                    stepIndex := 8; // Cycle complete, stay here
                END_IF;
        END_CASE;

    ELSIF ContinuousMode THEN
        // Continuous mode: run through all steps automatically, restart at end
        CASE stepIndex OF
            0:
                MoveDown := NOT DownLimitSwitch;
                IF DownLimitSwitch THEN
                    stepIndex := 1;
                END_IF;
            1:
                ActivateGrip := NOT GripLimitSwitch;
                IF GripLimitSwitch THEN
                    stepIndex := 2;
                END_IF;
            2:
                MoveUp := NOT UpLimitSwitch;
                IF UpLimitSwitch THEN
                    stepIndex := 3;
                END_IF;
            3:
                MoveRight := NOT RightLimitSwitch;
                IF RightLimitSwitch THEN
                    stepIndex := 4;
                END_IF;
            4:
                MoveDown := NOT DownLimitSwitch;
                IF DownLimitSwitch THEN
                    stepIndex := 5;
                END_IF;
            5:
                ActivateRelease := NOT ReleaseLimitSwitch;
                IF ReleaseLimitSwitch THEN
                    stepIndex := 6;
                END_IF;
            6:
                MoveUp := NOT UpLimitSwitch;
                IF UpLimitSwitch THEN
                    stepIndex := 7;
                END_IF;
            7:
                MoveLeft := NOT LeftLimitSwitch;
                IF LeftLimitSwitch THEN
                    stepIndex := 0; // Restart cycle
                END_IF;
        END_CASE;

    ELSIF ManualMode THEN
        // Manual mode: direct button control with limit switch protection
        MoveDown := DownButton AND NOT DownLimitSwitch;
        MoveUp := UpButton AND NOT UpLimitSwitch;
        MoveLeft := LeftButton AND NOT LeftLimitSwitch;
        MoveRight := RightButton AND NOT RightLimitSwitch;
        ActivateGrip := GripButton AND NOT GripLimitSwitch;
        ActivateRelease := ReleaseButton AND NOT ReleaseLimitSwitch;
    END_IF;

END_FUNCTION_BLOCK

(* ---- public-hard-05.patch_base_03.st ---- *)
(* ENGINEERING_CONTRACT - Mechanical Arm Control
 * =============================================================================
 * Mode Selection: Caller ensures exactly one mode active; emergency stop has highest priority.
 *
 * Output State Table:
 * | Output          | Activation                              | Retention                     | Reset                        | Priority    |
 * |-----------------|-----------------------------------------|-------------------------------|--------------------------------|-------------|
 * | MoveDown        | Manual:DownButton AND NOT DownLimitSwitch| Manual:button hold; Auto:step | EmergencyStop, step change   | Physical dir |
 * |                 | Auto: current step = down step           | Auto: hold until limit        | button release (manual)       | rule applies |
 * | MoveUp          | Manual:UpButton AND NOT UpLimitSwitch    | Manual:button hold; Auto:step | EmergencyStop, step change   | Physical dir |
 * |                 | Auto: current step = up step             | Auto: hold until limit        | button release (manual)       | rule applies |
 * | MoveLeft        | Manual:LeftButton AND NOT LeftLimitSwitch| Manual:button hold; Auto:step | EmergencyStop, step change   | Physical dir |
 * |                 | Auto: current step = left step           | Auto: hold until limit        | button release (manual)       | rule applies |
 * | MoveRight       | Manual:RightButton AND NOT RightLimitSwitch| Manual:button hold; Auto:step| EmergencyStop, step change   | Physical dir |
 * |                 | Auto: current step = right step          | Auto: hold until limit        | button release (manual)       | rule applies |
 * | ActivateGrip    | Manual:GripButton AND NOT GripLimitSwitch| Manual:button hold; Auto:step | EmergencyStop, step change   | N/A         |
 * |                 | Auto: grip step, hold until GripLimitSwitch| Auto: hold until limit       | button release (manual)       |             |
 * | ActivateRelease | Manual:ReleaseButton AND NOT ReleaseLimitSwitch| Manual:button hold; Auto:step| EmergencyStop, step change  | N/A         |
 * |                 | Auto: release step, hold until ReleaseLimitSwitch| Auto: hold until limit    | button release (manual)       |             |
 *
 * Sequence (8 steps, single cycle and continuous modes):
 *   0: Down -> 1: Grip -> 2: Up -> 3: Right -> 4: Down -> 5: Release -> 6: Up -> 7: Left -> (repeat)
 *
 * Single step mode: Same 8-step sequence, advancing one step per Start rising edge.
 * Single cycle mode: Executes all 8 steps, stops at stepIndex=8.
 * Continuous mode: Executes all 8 steps, returns to stepIndex=0 when complete.
 *
 * Units: Limit switches TRUE=at position (normally-open, closed at position).
 * Boundary: stepIndex ∈ [0..8]; 8 = cycle complete state for single cycle mode.
 * Same-scan: Final output evaluated from current stepIndex and limit switches per scan.
 *
 * Contract PUB clauses: PUB001-PUB020 define all behavior above.
 *)

FUNCTION_BLOCK ArmController
VAR_INPUT
    ManualMode : BOOL;
    SingleStepMode : BOOL;
    SingleCycleMode : BOOL;
    ContinuousMode : BOOL;
    EmergencyStop : BOOL;
    Start : BOOL;
    DownButton : BOOL;
    UpButton : BOOL;
    LeftButton : BOOL;
    RightButton : BOOL;
    GripButton : BOOL;
    ReleaseButton : BOOL;
    DownLimitSwitch : BOOL;
    UpLimitSwitch : BOOL;
    LeftLimitSwitch : BOOL;
    RightLimitSwitch : BOOL;
    GripLimitSwitch : BOOL;
    ReleaseLimitSwitch : BOOL;
END_VAR
VAR_OUTPUT
    MoveDown : BOOL;
    MoveUp : BOOL;
    MoveLeft : BOOL;
    MoveRight : BOOL;
    ActivateGrip : BOOL;
    ActivateRelease : BOOL;
END_VAR
VAR
    stepIndex : INT := 0;         // Current step in sequence (0-7), 8 = single cycle complete
    startButtonPrev : BOOL := FALSE; // Rising edge detection for Start button
    tmpRisingEdge : BOOL;
END_VAR

(* CONTRACT_RULES
[
  {"kind": "hold_until_reset", "output": "MoveDown", "set_input": "DownButton", "reset_input": null},
  {"kind": "hold_until_reset", "output": "MoveUp", "set_input": "UpButton", "reset_input": null},
  {"kind": "hold_until_reset", "output": "MoveLeft", "set_input": "LeftButton", "reset_input": null},
  {"kind": "hold_until_reset", "output": "MoveRight", "set_input": "RightButton", "reset_input": null},
  {"kind": "hold_until_reset", "output": "ActivateGrip", "set_input": "GripButton", "reset_input": null},
  {"kind": "hold_until_reset", "output": "ActivateRelease", "set_input": "ReleaseButton", "reset_input": null}
]
*)

    // Emergency stop has highest priority - stops all outputs
    IF EmergencyStop = FALSE THEN
        MoveDown := FALSE;
        MoveUp := FALSE;
        MoveLeft := FALSE;
        MoveRight := FALSE;
        ActivateGrip := FALSE;
        ActivateRelease := FALSE;
    ELSIF SingleStepMode THEN
        // Detect rising edge on Start button
        tmpRisingEdge := Start AND NOT startButtonPrev;
        startButtonPrev := Start;

        IF tmpRisingEdge THEN
            stepIndex := stepIndex + 1;
            IF stepIndex > 7 THEN
                stepIndex := 0;
            END_IF;
        END_IF;

        // Execute current step
        CASE stepIndex OF
            0: // Down
                MoveDown := TRUE;
                IF DownLimitSwitch THEN
                    stepIndex := 1;
                END_IF;
            1: // Grip
                ActivateGrip := TRUE;
                IF GripLimitSwitch THEN
                    stepIndex := 2;
                END_IF;
            2: // Up
                MoveUp := TRUE;
                IF UpLimitSwitch THEN
                    stepIndex := 3;
                END_IF;
            3: // Right
                MoveRight := TRUE;
                IF RightLimitSwitch THEN
                    stepIndex := 4;
                END_IF;
            4: // Down (second descent)
                MoveDown := TRUE;
                IF DownLimitSwitch THEN
                    stepIndex := 5;
                END_IF;
            5: // Release
                ActivateRelease := TRUE;
                IF ReleaseLimitSwitch THEN
                    stepIndex := 6;
                END_IF;
            6: // Up (second ascent)
                MoveUp := TRUE;
                IF UpLimitSwitch THEN
                    stepIndex := 7;
                END_IF;
            7: // Left (return to start)
                MoveLeft := TRUE;
                IF LeftLimitSwitch THEN
                    stepIndex := 0;
                END_IF;
        END_CASE;

    ELSIF SingleCycleMode THEN
        // Single cycle mode: run through all steps automatically, stop at end
        CASE stepIndex OF
            0:
                MoveDown := NOT DownLimitSwitch;
                IF DownLimitSwitch THEN
                    stepIndex := 1;
                END_IF;
            1:
                ActivateGrip := NOT GripLimitSwitch;
                IF GripLimitSwitch THEN
                    stepIndex := 2;
                END_IF;
            2:
                MoveUp := NOT UpLimitSwitch;
                IF UpLimitSwitch THEN
                    stepIndex := 3;
                END_IF;
            3:
                MoveRight := NOT RightLimitSwitch;
                IF RightLimitSwitch THEN
                    stepIndex := 4;
                END_IF;
            4:
                MoveDown := NOT DownLimitSwitch;
                IF DownLimitSwitch THEN
                    stepIndex := 5;
                END_IF;
            5:
                ActivateRelease := NOT ReleaseLimitSwitch;
                IF ReleaseLimitSwitch THEN
                    stepIndex := 6;
                END_IF;
            6:
                MoveUp := NOT UpLimitSwitch;
                IF UpLimitSwitch THEN
                    stepIndex := 7;
                END_IF;
            7:
                MoveLeft := NOT LeftLimitSwitch;
                IF LeftLimitSwitch THEN
                    stepIndex := 8; // Cycle complete, stay here
                END_IF;
        END_CASE;

    ELSIF ContinuousMode THEN
        // Continuous mode: run through all steps automatically, restart at end
        CASE stepIndex OF
            0:
                MoveDown := NOT DownLimitSwitch;
                IF DownLimitSwitch THEN
                    stepIndex := 1;
                END_IF;
            1:
                ActivateGrip := NOT GripLimitSwitch;
                IF GripLimitSwitch THEN
                    stepIndex := 2;
                END_IF;
            2:
                MoveUp := NOT UpLimitSwitch;
                IF UpLimitSwitch THEN
                    stepIndex := 3;
                END_IF;
            3:
                MoveRight := NOT RightLimitSwitch;
                IF RightLimitSwitch THEN
                    stepIndex := 4;
                END_IF;
            4:
                MoveDown := NOT DownLimitSwitch;
                IF DownLimitSwitch THEN
                    stepIndex := 5;
                END_IF;
            5:
                ActivateRelease := NOT ReleaseLimitSwitch;
                IF ReleaseLimitSwitch THEN
                    stepIndex := 6;
                END_IF;
            6:
                MoveUp := NOT UpLimitSwitch;
                IF UpLimitSwitch THEN
                    stepIndex := 7;
                END_IF;
            7:
                MoveLeft := NOT LeftLimitSwitch;
                IF LeftLimitSwitch THEN
                    stepIndex := 0; // Restart cycle
                END_IF;
        END_CASE;

    ELSIF ManualMode THEN
        // Manual mode: direct button control with limit switch protection
        MoveDown := DownButton AND NOT DownLimitSwitch;
        MoveUp := UpButton AND NOT UpLimitSwitch;
        MoveLeft := LeftButton AND NOT LeftLimitSwitch;
        MoveRight := RightButton AND NOT RightLimitSwitch;
        ActivateGrip := GripButton AND NOT GripLimitSwitch;
        ActivateRelease := ReleaseButton AND NOT ReleaseLimitSwitch;
    END_IF;

END_FUNCTION_BLOCK

(* ---- public-hard-05.patch_base_04.st ---- *)
(* ENGINEERING_CONTRACT - Mechanical Arm Control
 * =============================================================================
 * Mode Selection: Caller ensures exactly one mode active; emergency stop has highest priority.
 *
 * Output State Table:
 * | Output          | Activation                              | Retention                     | Reset                        | Priority    |
 * |-----------------|-----------------------------------------|-------------------------------|--------------------------------|-------------|
 * | MoveDown        | Manual:DownButton AND NOT DownLimitSwitch| Manual:button hold; Auto:step | EmergencyStop, step change   | Physical dir |
 * |                 | Auto: current step = down step           | Auto: hold until limit        | button release (manual)       | rule applies |
 * | MoveUp          | Manual:UpButton AND NOT UpLimitSwitch    | Manual:button hold; Auto:step | EmergencyStop, step change   | Physical dir |
 * |                 | Auto: current step = up step             | Auto: hold until limit        | button release (manual)       | rule applies |
 * | MoveLeft        | Manual:LeftButton AND NOT LeftLimitSwitch| Manual:button hold; Auto:step | EmergencyStop, step change   | Physical dir |
 * |                 | Auto: current step = left step           | Auto: hold until limit        | button release (manual)       | rule applies |
 * | MoveRight       | Manual:RightButton AND NOT RightLimitSwitch| Manual:button hold; Auto:step| EmergencyStop, step change   | Physical dir |
 * |                 | Auto: current step = right step          | Auto: hold until limit        | button release (manual)       | rule applies |
 * | ActivateGrip    | Manual:GripButton AND NOT GripLimitSwitch| Manual:button hold; Auto:step | EmergencyStop, step change   | N/A         |
 * |                 | Auto: grip step, hold until GripLimitSwitch| Auto: hold until limit       | button release (manual)       |             |
 * | ActivateRelease | Manual:ReleaseButton AND NOT ReleaseLimitSwitch| Manual:button hold; Auto:step| EmergencyStop, step change  | N/A         |
 * |                 | Auto: release step, hold until ReleaseLimitSwitch| Auto: hold until limit    | button release (manual)       |             |
 *
 * Sequence (8 steps, single cycle and continuous modes):
 *   0: Down -> 1: Grip -> 2: Up -> 3: Right -> 4: Down -> 5: Release -> 6: Up -> 7: Left -> (repeat)
 *
 * Single step mode: Same 8-step sequence, advancing one step per Start rising edge.
 * Single cycle mode: Executes all 8 steps, stops at stepIndex=8.
 * Continuous mode: Executes all 8 steps, returns to stepIndex=0 when complete.
 *
 * Units: Limit switches TRUE=at position (normally-open, closed at position).
 * Boundary: stepIndex ∈ [0..8]; 8 = cycle complete state for single cycle mode.
 * Same-scan: Final output evaluated from current stepIndex and limit switches per scan.
 *
 * Contract PUB clauses: PUB001-PUB020 define all behavior above.
 *)

FUNCTION_BLOCK ArmController
VAR_INPUT
    ManualMode : BOOL;
    SingleStepMode : BOOL;
    SingleCycleMode : BOOL;
    ContinuousMode : BOOL;
    EmergencyStop : BOOL;
    Start : BOOL;
    DownButton : BOOL;
    UpButton : BOOL;
    LeftButton : BOOL;
    RightButton : BOOL;
    GripButton : BOOL;
    ReleaseButton : BOOL;
    DownLimitSwitch : BOOL;
    UpLimitSwitch : BOOL;
    LeftLimitSwitch : BOOL;
    RightLimitSwitch : BOOL;
    GripLimitSwitch : BOOL;
    ReleaseLimitSwitch : BOOL;
END_VAR
VAR_OUTPUT
    MoveDown : BOOL;
    MoveUp : BOOL;
    MoveLeft : BOOL;
    MoveRight : BOOL;
    ActivateGrip : BOOL;
    ActivateRelease : BOOL;
END_VAR
VAR
    stepIndex : INT := 0;         // Current step in sequence (0-7), 8 = single cycle complete
    startButtonPrev : BOOL := FALSE; // Rising edge detection for Start button
    tmpRisingEdge : BOOL;
END_VAR

(* CONTRACT_RULES
[
  {"kind": "hold_until_reset", "output": "MoveDown", "set_input": "DownButton", "reset_input": null},
  {"kind": "hold_until_reset", "output": "MoveUp", "set_input": "UpButton", "reset_input": null},
  {"kind": "hold_until_reset", "output": "MoveLeft", "set_input": "LeftButton", "reset_input": null},
  {"kind": "hold_until_reset", "output": "MoveRight", "set_input": "RightButton", "reset_input": null},
  {"kind": "hold_until_reset", "output": "ActivateGrip", "set_input": "GripButton", "reset_input": null},
  {"kind": "hold_until_reset", "output": "ActivateRelease", "set_input": "ReleaseButton", "reset_input": null}
]
*)

    // Emergency stop has highest priority - stops all outputs
    IF EmergencyStop = FALSE THEN
        MoveDown := FALSE;
        MoveUp := FALSE;
        MoveLeft := FALSE;
        MoveRight := FALSE;
        ActivateGrip := FALSE;
        ActivateRelease := FALSE;
    ELSIF SingleStepMode THEN
        // Detect rising edge on Start button
        tmpRisingEdge := Start AND NOT startButtonPrev;
        startButtonPrev := Start;

        IF tmpRisingEdge THEN
            stepIndex := stepIndex + 1;
            IF stepIndex > 7 THEN
                stepIndex := 0;
            END_IF;
        END_IF;

        // Execute current step
        CASE stepIndex OF
            0: // Down
                MoveDown := TRUE;
                IF DownLimitSwitch THEN
                    stepIndex := 1;
                END_IF;
            1: // Grip
                ActivateGrip := TRUE;
                IF GripLimitSwitch THEN
                    stepIndex := 2;
                END_IF;
            2: // Up
                MoveUp := TRUE;
                IF UpLimitSwitch THEN
                    stepIndex := 3;
                END_IF;
            3: // Right
                MoveRight := TRUE;
                IF RightLimitSwitch THEN
                    stepIndex := 4;
                END_IF;
            4: // Down (second descent)
                MoveDown := TRUE;
                IF DownLimitSwitch THEN
                    stepIndex := 5;
                END_IF;
            5: // Release
                ActivateRelease := TRUE;
                IF ReleaseLimitSwitch THEN
                    stepIndex := 6;
                END_IF;
            6: // Up (second ascent)
                MoveUp := TRUE;
                IF UpLimitSwitch THEN
                    stepIndex := 7;
                END_IF;
            7: // Left (return to start)
                MoveLeft := TRUE;
                IF LeftLimitSwitch THEN
                    stepIndex := 0;
                END_IF;
        END_CASE;

    ELSIF SingleCycleMode THEN
        // Single cycle mode: run through all steps automatically, stop at end
        CASE stepIndex OF
            0:
                MoveDown := NOT DownLimitSwitch;
                IF DownLimitSwitch THEN
                    stepIndex := 1;
                END_IF;
            1:
                ActivateGrip := NOT GripLimitSwitch;
                IF GripLimitSwitch THEN
                    stepIndex := 2;
                END_IF;
            2:
                MoveUp := NOT UpLimitSwitch;
                IF UpLimitSwitch THEN
                    stepIndex := 3;
                END_IF;
            3:
                MoveRight := NOT RightLimitSwitch;
                IF RightLimitSwitch THEN
                    stepIndex := 4;
                END_IF;
            4:
                MoveDown := NOT DownLimitSwitch;
                IF DownLimitSwitch THEN
                    stepIndex := 5;
                END_IF;
            5:
                ActivateRelease := NOT ReleaseLimitSwitch;
                IF ReleaseLimitSwitch THEN
                    stepIndex := 6;
                END_IF;
            6:
                MoveUp := NOT UpLimitSwitch;
                IF UpLimitSwitch THEN
                    stepIndex := 7;
                END_IF;
            7:
                MoveLeft := NOT LeftLimitSwitch;
                IF LeftLimitSwitch THEN
                    stepIndex := 8; // Cycle complete, stay here
                END_IF;
        END_CASE;

    ELSIF ContinuousMode THEN
        // Continuous mode: run through all steps automatically, restart at end
        CASE stepIndex OF
            0:
                MoveDown := NOT DownLimitSwitch;
                IF DownLimitSwitch THEN
                    stepIndex := 1;
                END_IF;
            1:
                ActivateGrip := NOT GripLimitSwitch;
                IF GripLimitSwitch THEN
                    stepIndex := 2;
                END_IF;
            2:
                MoveUp := NOT UpLimitSwitch;
                IF UpLimitSwitch THEN
                    stepIndex := 3;
                END_IF;
            3:
                MoveRight := NOT RightLimitSwitch;
                IF RightLimitSwitch THEN
                    stepIndex := 4;
                END_IF;
            4:
                MoveDown := NOT DownLimitSwitch;
                IF DownLimitSwitch THEN
                    stepIndex := 5;
                END_IF;
            5:
                ActivateRelease := NOT ReleaseLimitSwitch;
                IF ReleaseLimitSwitch THEN
                    stepIndex := 6;
                END_IF;
            6:
                MoveUp := NOT UpLimitSwitch;
                IF UpLimitSwitch THEN
                    stepIndex := 7;
                END_IF;
            7:
                MoveLeft := NOT LeftLimitSwitch;
                IF LeftLimitSwitch THEN
                    stepIndex := 0; // Restart cycle
                END_IF;
        END_CASE;

    ELSIF ManualMode THEN
        // Manual mode: direct button control with limit switch protection
        MoveDown := DownButton AND NOT DownLimitSwitch;
        MoveUp := UpButton AND NOT UpLimitSwitch;
        MoveLeft := LeftButton AND NOT LeftLimitSwitch;
        MoveRight := RightButton AND NOT RightLimitSwitch;
        ActivateGrip := GripButton AND NOT GripLimitSwitch;
        ActivateRelease := ReleaseButton AND NOT ReleaseLimitSwitch;
    END_IF;

END_FUNCTION_BLOCK
